//{attribute 'qualified_only'}
VAR_GLOBAL
	i_EL			AT %I*	: ARRAY[1..27] 		OF ST_EL18x9;
	q_EL			AT %Q*	: ARRAY[1..11] 		OF ST_EL28x9;
	ai_EL			AT %I*	: ARRAY[1..6] 		OF ST_EL3xx8;
	aq_EL			AT %Q*	: ARRAY[1..1] 		OF ST_EL4xx8;

	
	q_Manifold1 	AT %Q*	: ARRAY[1..24] 		OF ST_VTUG;
	q_Manifold2 	AT %Q*	: ARRAY[1..24] 		OF ST_VTUG;
	q_Manifold3 	AT %Q*	: ARRAY[1..24] 		OF ST_VTUG;

	Nidec					: ARRAY[0..E_Pump_List.last] 		OF ST_Nidec;

	
	arSafe			: ARRAY[1..1] OF ST_TwinSAFE;
	bStateSafe		: BOOL;
	bStateSafe_ES1	: BOOL;
	bStateSafe_ES2	: BOOL;
	bStateSafe_ES3	: BOOL;
	bStateSafe_ES4	: BOOL;
	
	fbScaleFactor: ARRAY[0..E_ASense_Name.last] 		OF FB_ScaleFactor;
	
	//Anybus Communicator (Box 40), 128 bytes each direction, decoded in g_Anybus.fbAnybus
	Anybus_Inputs_Raw  AT %I* : ARRAY [0..127] OF BYTE;
    Anybus_Outputs_Raw AT %Q* : ARRAY [0..127] OF BYTE;
	Anybus_WcState     AT %I* : BOOL;	//Box 40 WcState, TRUE = process data not valid (also when not in OP)

	
END_VAR

(* stored: Version 1.1.0.1, ProductVersion 3.1.4026.20
   GVL gIO: Id {d074f1fc-f55a-4f30-b093-dc5be34740ab} *)
